(* IEC 61131-3 sources: Caravan/Archiv/12-04-19/Stations/Terminal/HMI/Network/WEATHER_WeatherForecast, 1 file *)

(* ---- ONE_WEATHER_WeatherForecast_Table.st ---- *)
#define OBJECTS_CONFIG

//Define part of class _WeatherForecast
//=====================================================================================================================

#define WEATHERFC_DEF_URL_P1  "http://api.openweathermap.org/data/2.5/forecast?"   // URL Default part 1
#define WEATHERFC_DEF_URL_EXT "&units=metric&mode=xml"                             // URL Default extensions

#define WEATHERFC_XmlFile     "WeatherForecast.xml"   // Name of the XML-file

#define WEATHERFC_XmlEntries  40                      // Number of entries in the weather-xml (5 days * 8 entries/day)

#define NEW_DATA_IN_PROCESS    99                     // staus "new data will be processed"
#define HTTP_REQUEST_OK       200                     // http return code "everything ok"

//=====================================================================================================================
#include <.\lsl_st_httpclient.h>

FUNCTION GLOBAL TAB ONE_WEATHER_WeatherForecast
-1$UINT, 0$UINT,
0$UINT, 0$UINT,

10$UDINT,
TO_UDINT(2980745877), "_MyIO", 0$UINT, 3$UINT, 0$UINT,
TO_UDINT(3839744317), "_WeatherForecast", 1$UINT, 1$UINT, 1$UINT,
TO_UDINT(428324901), "_WindIndicator", 1$UINT, 0$UINT, 1$UINT,
TO_UDINT(3727258101), "_XMLReader", 1$UINT, 4$UINT, 1$UINT,
TO_UDINT(2131172539), "_XMLStructCreator", 1$UINT, 2$UINT, 1$UINT,
TO_UDINT(2225119864), "MerkerEx", 1$UINT, 21$UINT, 0$UINT,
TO_UDINT(933570811), "RAMex", 1$UINT, 17$UINT, 15$UINT,
TO_UDINT(2898603620), "StringInternal", 1$UINT, 82$UINT, 0$UINT,
TO_UDINT(2408581120), "StringRAM", 1$UINT, 10$UINT, 15$UINT,
TO_UDINT(3232495061), "VirtualBaseInit", 1$UINT, 3$UINT, 0$UINT,

_NO_ATTR, TO_UDINT(3679485567), "_WEATHERFORECAST1",

_NO_ATTR, TO_UDINT(3368139848), "_WINDINDICATOR1",

_NO_ATTR, TO_UDINT(1322631253), "_XMLREADER1",

1$UINT, TO_UDINT(4272249074), "_XMLREADER1\STRUCTCREATOR",

1$UINT, TO_UDINT(2164056838), "_WEATHERFORECAST1\STR_DAY1_DD_MM\DATABUFFER",
1$UINT, TO_UDINT(1786396260), "_WEATHERFORECAST1\STR_DAY2_DD_MM\DATABUFFER",
1$UINT, TO_UDINT(2234026117), "_WEATHERFORECAST1\STR_DAY3_DD_MM\DATABUFFER",
1$UINT, TO_UDINT(1678148321), "_WEATHERFORECAST1\STR_DAY4_DD_MM\DATABUFFER",
1$UINT, TO_UDINT(2337551360), "_WEATHERFORECAST1\STR_DAY5_DD_MM\DATABUFFER",
1$UINT, TO_UDINT(2939021694), "_WEATHERFORECAST1\STR_LASTLOCATIONNAME\DATABUFFER",
1$UINT, TO_UDINT(3127945444), "_WEATHERFORECAST1\STR_PROXYADDRESS\DATABUFFER",
1$UINT, TO_UDINT(298110734), "_WEATHERFORECAST1\STR_PROXYPASSWORD\DATABUFFER",
1$UINT, TO_UDINT(274360433), "_WEATHERFORECAST1\STR_PROXYPORT\DATABUFFER",
1$UINT, TO_UDINT(1238597337), "_WEATHERFORECAST1\STR_PROXYUSER\DATABUFFER",
1$UINT, TO_UDINT(3526506352), "_WEATHERFORECAST1\STR_WEATHERLOCCOUNTRY\DATABUFFER",
1$UINT, TO_UDINT(3122055684), "_WEATHERFORECAST1\STR_WEATHERLOCID\DATABUFFER",
1$UINT, TO_UDINT(1698372815), "_WEATHERFORECAST1\STR_WEATHERLOCNAME\DATABUFFER",
1$UINT, TO_UDINT(3270495593), "_WEATHERFORECAST1\STR_WEATHERURL\DATABUFFER",
1$UINT, TO_UDINT(246742247), "_WEATHERFORECAST1\STR_WEATHERUSERID\DATABUFFER",

1$UINT, TO_UDINT(2519093562), "_WEATHERFORECAST1\STR_DAY1_DD_MM",
1$UINT, TO_UDINT(2815314855), "_WEATHERFORECAST1\STR_DAY2_DD_MM",
1$UINT, TO_UDINT(28917779), "_WEATHERFORECAST1\STR_DAY3_DD_MM",
1$UINT, TO_UDINT(3290332829), "_WEATHERFORECAST1\STR_DAY4_DD_MM",
1$UINT, TO_UDINT(1651078441), "_WEATHERFORECAST1\STR_DAY5_DD_MM",
1$UINT, TO_UDINT(3331481044), "_WEATHERFORECAST1\STR_LASTLOCATIONNAME",
1$UINT, TO_UDINT(2090602944), "_WEATHERFORECAST1\STR_PROXYADDRESS",
1$UINT, TO_UDINT(252101989), "_WEATHERFORECAST1\STR_PROXYPASSWORD",
1$UINT, TO_UDINT(2245335798), "_WEATHERFORECAST1\STR_PROXYPORT",
1$UINT, TO_UDINT(1272418675), "_WEATHERFORECAST1\STR_PROXYUSER",
1$UINT, TO_UDINT(2168826918), "_WEATHERFORECAST1\STR_WEATHERLOCCOUNTRY",
1$UINT, TO_UDINT(1133894061), "_WEATHERFORECAST1\STR_WEATHERLOCID",
1$UINT, TO_UDINT(2097317819), "_WEATHERFORECAST1\STR_WEATHERLOCNAME",
1$UINT, TO_UDINT(2424888079), "_WEATHERFORECAST1\STR_WEATHERURL",
1$UINT, TO_UDINT(183002200), "_WEATHERFORECAST1\STR_WEATHERUSERID",

//Internal connections
0$UDINT,
31$UDINT,
TO_UDINT(0), "Str_WeatherURL", TO_UDINT(32),
TO_UDINT(0), "Str_ProxyPort", TO_UDINT(27),
TO_UDINT(0), "Str_ProxyUser", TO_UDINT(28),
TO_UDINT(0), "Str_ProxyPassword", TO_UDINT(26),
TO_UDINT(0), "Str_WeatherUserID", TO_UDINT(33),
TO_UDINT(0), "Str_WeatherLocName", TO_UDINT(31),
TO_UDINT(0), "Str_WeatherLocCountry", TO_UDINT(29),
TO_UDINT(0), "Str_WeatherLocID", TO_UDINT(30),
TO_UDINT(0), "Str_ProxyAddress", TO_UDINT(25),
TO_UDINT(0), "Str_Day1_DD_MM", TO_UDINT(19),
TO_UDINT(0), "Str_Day2_DD_MM", TO_UDINT(20),
TO_UDINT(0), "Str_Day3_DD_MM", TO_UDINT(21),
TO_UDINT(0), "Str_Day4_DD_MM", TO_UDINT(22),
TO_UDINT(0), "Str_Day5_DD_MM", TO_UDINT(23),
TO_UDINT(0), "Str_LastLocationName", TO_UDINT(24),
TO_UDINT(2), "StructCreator", TO_UDINT(3),
TO_UDINT(19), "DataBuffer", TO_UDINT(4),
TO_UDINT(20), "DataBuffer", TO_UDINT(5),
TO_UDINT(21), "DataBuffer", TO_UDINT(6),
TO_UDINT(22), "DataBuffer", TO_UDINT(7),
TO_UDINT(23), "DataBuffer", TO_UDINT(8),
TO_UDINT(24), "DataBuffer", TO_UDINT(9),
TO_UDINT(25), "DataBuffer", TO_UDINT(10),
TO_UDINT(26), "DataBuffer", TO_UDINT(11),
TO_UDINT(27), "DataBuffer", TO_UDINT(12),
TO_UDINT(28), "DataBuffer", TO_UDINT(13),
TO_UDINT(29), "DataBuffer", TO_UDINT(14),
TO_UDINT(30), "DataBuffer", TO_UDINT(15),
TO_UDINT(31), "DataBuffer", TO_UDINT(16),
TO_UDINT(32), "DataBuffer", TO_UDINT(17),
TO_UDINT(33), "DataBuffer", TO_UDINT(18),
0$UDINT,
17$UDINT,
TO_UDINT(0), "_XMLReader", TO_UDINT(2), "ClassSvr",
TO_UDINT(1), "WindDirection", TO_UDINT(0), "Day1WindDegree",
TO_UDINT(19), "DataBuffer", TO_UDINT(4), "m_udLength",
TO_UDINT(20), "DataBuffer", TO_UDINT(5), "m_udLength",
TO_UDINT(21), "DataBuffer", TO_UDINT(6), "m_udLength",
TO_UDINT(22), "DataBuffer", TO_UDINT(7), "m_udLength",
TO_UDINT(23), "DataBuffer", TO_UDINT(8), "m_udLength",
TO_UDINT(24), "DataBuffer", TO_UDINT(9), "m_udLength",
TO_UDINT(25), "DataBuffer", TO_UDINT(10), "m_udLength",
TO_UDINT(26), "DataBuffer", TO_UDINT(11), "m_udLength",
TO_UDINT(27), "DataBuffer", TO_UDINT(12), "m_udLength",
TO_UDINT(28), "DataBuffer", TO_UDINT(13), "m_udLength",
TO_UDINT(29), "DataBuffer", TO_UDINT(14), "m_udLength",
TO_UDINT(30), "DataBuffer", TO_UDINT(15), "m_udLength",
TO_UDINT(31), "DataBuffer", TO_UDINT(16), "m_udLength",
TO_UDINT(32), "DataBuffer", TO_UDINT(17), "m_udLength",
TO_UDINT(33), "DataBuffer", TO_UDINT(18), "m_udLength",

//Initialization values
0$UDINT,
32$UDINT,
TO_UDINT(0), "AutoUpdate", TO_UDINT(15),//|WEATHER_WeatherForecast._WeatherForecast1.AutoUpdate;
TO_UDINT(0), "UTC_Offset", TO_UDINT(0),//|WEATHER_WeatherForecast._WeatherForecast1.UTC_Offset;
TO_UDINT(4), "ThreadSafe", TO_UDINT(0),//|WEATHER_WeatherForecast.Str_Day1_DD_MM\_WeatherForecast1\DataBuffer.ThreadSafe;
TO_UDINT(5), "ThreadSafe", TO_UDINT(0),//|WEATHER_WeatherForecast.Str_Day2_DD_MM\_WeatherForecast1\DataBuffer.ThreadSafe;
TO_UDINT(6), "ThreadSafe", TO_UDINT(0),//|WEATHER_WeatherForecast.Str_Day3_DD_MM\_WeatherForecast1\DataBuffer.ThreadSafe;
TO_UDINT(7), "ThreadSafe", TO_UDINT(0),//|WEATHER_WeatherForecast.Str_Day4_DD_MM\_WeatherForecast1\DataBuffer.ThreadSafe;
TO_UDINT(8), "ThreadSafe", TO_UDINT(0),//|WEATHER_WeatherForecast.Str_Day5_DD_MM\_WeatherForecast1\DataBuffer.ThreadSafe;
TO_UDINT(9), "ThreadSafe", TO_UDINT(0),//|WEATHER_WeatherForecast.Str_LastLocationName\_WeatherForecast1\DataBuffer.ThreadSafe;
TO_UDINT(10), "ThreadSafe", TO_UDINT(0),//|WEATHER_WeatherForecast.Str_ProxyAddress\_WeatherForecast1\DataBuffer.ThreadSafe;
TO_UDINT(11), "ThreadSafe", TO_UDINT(0),//|WEATHER_WeatherForecast.Str_ProxyPassword\_WeatherForecast1\DataBuffer.ThreadSafe;
TO_UDINT(12), "ThreadSafe", TO_UDINT(0),//|WEATHER_WeatherForecast.Str_ProxyPort\_WeatherForecast1\DataBuffer.ThreadSafe;
TO_UDINT(13), "ThreadSafe", TO_UDINT(0),//|WEATHER_WeatherForecast.Str_ProxyUser\_WeatherForecast1\DataBuffer.ThreadSafe;
TO_UDINT(14), "ThreadSafe", TO_UDINT(0),//|WEATHER_WeatherForecast.Str_WeatherLocCountry\_WeatherForecast1\DataBuffer.ThreadSafe;
TO_UDINT(15), "ThreadSafe", TO_UDINT(0),//|WEATHER_WeatherForecast.Str_WeatherLocID\_WeatherForecast1\DataBuffer.ThreadSafe;
TO_UDINT(16), "ThreadSafe", TO_UDINT(0),//|WEATHER_WeatherForecast.Str_WeatherLocName\_WeatherForecast1\DataBuffer.ThreadSafe;
TO_UDINT(17), "ThreadSafe", TO_UDINT(0),//|WEATHER_WeatherForecast.Str_WeatherURL\_WeatherForecast1\DataBuffer.ThreadSafe;
TO_UDINT(18), "ThreadSafe", TO_UDINT(0),//|WEATHER_WeatherForecast.Str_WeatherUserID\_WeatherForecast1\DataBuffer.ThreadSafe;
TO_UDINT(19), "SingleRealloc", TO_UDINT(1),//|WEATHER_WeatherForecast._WeatherForecast1\Str_Day1_DD_MM.SingleRealloc;
TO_UDINT(20), "SingleRealloc", TO_UDINT(1),//|WEATHER_WeatherForecast._WeatherForecast1\Str_Day2_DD_MM.SingleRealloc;
TO_UDINT(21), "SingleRealloc", TO_UDINT(1),//|WEATHER_WeatherForecast._WeatherForecast1\Str_Day3_DD_MM.SingleRealloc;
TO_UDINT(22), "SingleRealloc", TO_UDINT(1),//|WEATHER_WeatherForecast._WeatherForecast1\Str_Day4_DD_MM.SingleRealloc;
TO_UDINT(23), "SingleRealloc", TO_UDINT(1),//|WEATHER_WeatherForecast._WeatherForecast1\Str_Day5_DD_MM.SingleRealloc;
TO_UDINT(24), "SingleRealloc", TO_UDINT(1),//|WEATHER_WeatherForecast._WeatherForecast1\Str_LastLocationName.SingleRealloc;
TO_UDINT(25), "SingleRealloc", TO_UDINT(1),//|WEATHER_WeatherForecast._WeatherForecast1\Str_ProxyAddress.SingleRealloc;
TO_UDINT(26), "SingleRealloc", TO_UDINT(1),//|WEATHER_WeatherForecast._WeatherForecast1\Str_ProxyPassword.SingleRealloc;
TO_UDINT(27), "SingleRealloc", TO_UDINT(1),//|WEATHER_WeatherForecast._WeatherForecast1\Str_ProxyPort.SingleRealloc;
TO_UDINT(28), "SingleRealloc", TO_UDINT(1),//|WEATHER_WeatherForecast._WeatherForecast1\Str_ProxyUser.SingleRealloc;
TO_UDINT(29), "SingleRealloc", TO_UDINT(1),//|WEATHER_WeatherForecast._WeatherForecast1\Str_WeatherLocCountry.SingleRealloc;
TO_UDINT(30), "SingleRealloc", TO_UDINT(1),//|WEATHER_WeatherForecast._WeatherForecast1\Str_WeatherLocID.SingleRealloc;
TO_UDINT(31), "SingleRealloc", TO_UDINT(1),//|WEATHER_WeatherForecast._WeatherForecast1\Str_WeatherLocName.SingleRealloc;
TO_UDINT(32), "SingleRealloc", TO_UDINT(1),//|WEATHER_WeatherForecast._WeatherForecast1\Str_WeatherURL.SingleRealloc;
TO_UDINT(33), "SingleRealloc", TO_UDINT(1),//|WEATHER_WeatherForecast._WeatherForecast1\Str_WeatherUserID.SingleRealloc;

//Symbolic initialization values
0$UDINT,
0$UDINT,

//Initialization of string values
0$UDINT,
0$UDINT,

//Configuration of tasks (RealTime, Cyclic, Background)
0$UDINT,
0$UDINT,

0$UDINT,
0$UDINT,

0$UDINT,
1$UDINT,
TO_UDINT(2), (100)$UDINT, 4194303$DINT, 	//_XMLREADER1

//External connections
0$UDINT,
2$UDINT,
TO_UDINT(0), "SDT_SysTime", C_DIR, TO_UDINT(3035062039), "SysDateTime","SysTime",
TO_UDINT(1), "Lse", C_DIR, TO_UDINT(299963966), "Lse","Lse",

//Magic internal connections
0$UDINT,
15$UDINT,
TO_UDINT(4), "UseFile", TO_UDINT(19), "UseFile",
TO_UDINT(5), "UseFile", TO_UDINT(20), "UseFile",
TO_UDINT(6), "UseFile", TO_UDINT(21), "UseFile",
TO_UDINT(7), "UseFile", TO_UDINT(22), "UseFile",
TO_UDINT(8), "UseFile", TO_UDINT(23), "UseFile",
TO_UDINT(9), "UseFile", TO_UDINT(24), "UseFile",
TO_UDINT(10), "UseFile", TO_UDINT(25), "UseFile",
TO_UDINT(11), "UseFile", TO_UDINT(26), "UseFile",
TO_UDINT(12), "UseFile", TO_UDINT(27), "UseFile",
TO_UDINT(13), "UseFile", TO_UDINT(28), "UseFile",
TO_UDINT(14), "UseFile", TO_UDINT(29), "UseFile",
TO_UDINT(15), "UseFile", TO_UDINT(30), "UseFile",
TO_UDINT(16), "UseFile", TO_UDINT(31), "UseFile",
TO_UDINT(17), "UseFile", TO_UDINT(32), "UseFile",
TO_UDINT(18), "UseFile", TO_UDINT(33), "UseFile",

//Configuration of timeslots of tasks (RealTime, Cyclic)
#ifdef __LSLLDR_TIMESLOTS__
0$UDINT,
0$UDINT,

0$UDINT,
0$UDINT,

#endif //__LSLLDR_TIMESLOTS__

//MultiMaster connections
#ifdef __LSLLDR_MULTIMASTER__
0$UDINT,
0$UDINT,
#endif //__LSLLDR_MULTIMASTER__

//Configuration for task ID (RealTime, CyclicTime)
#ifdef __LSLLDR_TASKID__
"\\\\TASKS2  "
0$UDINT,
0$UDINT,

0$UDINT,
0$UDINT,

0$UDINT,
1$UDINT,
(0)$UDINT, 	//_XMLREADER1

#endif //__LSLLDR_TASKID__

END_FUNCTION
